(* IEC 61131-3 sources: codesys-to-s7/tests/corpus/C2S7-SEM-SRRS/pos, 1 file *)

(* ---- input.st ---- *)
FUNCTION_BLOCK FB_Case
VAR
    f : SR;
    x : BOOL;
    y : BOOL;
END_VAR
f(SET1 := x, RESET := y);
END_FUNCTION_BLOCK
